{attribute 'qualified_only'}
{attribute 'strict'}
{attribute 'to_string'}
TYPE E_Default :
(
	eOptionA := 0,
	eOptionB,
	eOptionC
);
END_TYPE

(* stored: Version 1.1.0.1, ProductVersion 3.1.4026.19
   DUT E_Default: Id {2d47a2bf-eb95-4c07-bf02-b877cccbe14d} *)
